// TIA Portal V18 export
// export: Created 2026-11-25T00:00:00.0000000Z, ExportSetting WithDefaults
TagTable "Station"
  State :   ()
  Verdict :   ()
  NokCode :   ()
  FaultCode :   ()
  CntConsecNok :   ()
  Locked :   ()
  RigCheck :   ()
  CallOperator :   ()
  PartPresent :   ()
  TCycle :   ()
  CntTotal :   ()
  CntOk :   ()
  CntNok :   ()
  CntRejectConfirmed :   ()
  FpG1 :   ()
  FrG1 :   ()
  FMean :   ()
  FHyst :   ()
  FpG2 :   ()
  FPeak :   ()
  XPeak :   ()
  FStep :   ()
  XStop :   ()
  MeanLo :   ()
  MeanHi :   ()
  HystLo :   ()
  HystHi :   ()
  G2Lo :   ()
  G2Hi :   ()
  PeakFLo :   ()
  PeakFHi :   ()
  PeakXMin :   ()
  PeakXMax :   ()
  StepLo :   ()
  StopXLo :   ()
  StopXHi :   ()
